(* IEC 61131-3 sources: plc-hackathon-2026/work/dump/MyController/Plc Logic/Application/Profiles, 6 files *)

(* ---- Prof_EV.st ---- *)
// DATA_BLOCK "Prof_EV"
// NON_RETAIN
// EV sesije; indeks = punjac*300 + redni broj; Count = broj sesija po punjacu
   VAR_GLOBAL
      Count : Array[0..3] of Int;
      Arr : Array[0..1199] of DInt;
      Dep : Array[0..1199] of DInt;
      Energy : Array[0..1199] of Real;
   END_VAR

(* ---- Prof_FEC.st ---- *)
//DATA_BLOCK "Prof_FEC"
//{ S7_Optimized_Access := 'TRUE' }
//VERSION : 0.1
//NON_RETAIN
// Fiksna potrosnja [kW], Warehouse_15min_kW.csv
   VAR_GLOBAL
      Data : Array[0..35039] of Real;
   END_VAR

(* ---- Prof_FNE.st ---- *)
// DATA_BLOCK "Prof_FNE"
// { S7_Optimized_Access := 'TRUE' }
// VERSION : 0.1
// NON_RETAIN
// FNE [kW], PV_15min.csv (clip na 750 kW)
   VAR_GLOBAL
      Data : Array[0..35039] of Real;
   END_VAR

(* ---- Prof_PriceDA.st ---- *)
// DATA_BLOCK "Prof_PriceDA"
// NON_RETAIN
// Dan-unaprijed cijena [EUR/kWh], EL_prices_DA_2025.csv
   VAR_GLOBAL
      Data : Array[0..35039] of Real;
   END_VAR

(* ---- Prof_PriceTT.st ---- *)
// DATA_BLOCK "Prof_PriceTT"
// NON_RETAIN
// Dvotarifna cijena energije [EUR/kWh], EL_prices_Elektra_2025.csv
   VAR_GLOBAL
      Data : Array[0..35039] of Real;
   END_VAR

(* ---- Prof_VT.st ---- *)
// DATA_BLOCK "Prof_VT"
// NON_RETAIN
// TRUE = visa tarifa (izvedeno iz Elektra serije), koristi se za mrezarinu
   VAR_GLOBAL
      Data : Array[0..35039] of Bool;
   END_VAR
